(* IEC 61131-3 sources: PLC_I/plc/src/hardware, 9 files *)

(* ---- 全局变量_气缸IO映像.gvl.st ---- *)
(* 气缸物理 IO 映像。设备树把扩展输入/输出模块映射到本数组后，
   由 程序_气缸输入映射 / 程序_气缸输出映射 按工程表地址读写。
   容量：输入 112 点(7 WORD)，输出 56 点(4 WORD)。
   未映射时数组保持 0，模块在线位保持 FALSE，气缸许可因此关闭。 *)
VAR_GLOBAL CONSTANT
    ui气缸输入点数 : UINT := 112;
    ui气缸输出点数 : UINT := 56;
END_VAR
VAR_GLOBAL
    aw气缸输入映像 : ARRAY[0..6] OF WORD;
    aw气缸输出映像 : ARRAY[0..3] OF WORD;
    (* 真实模块诊断：由设备树/总线诊断赋值，不得用工程常量冒充。 *)
    b气缸输入模块在线 : BOOL;
    b气缸输出模块在线 : BOOL;
END_VAR

(* ---- 全局变量_气缸工程.gvl.st ---- *)
(* 唯一气缸工程配置：一缸一行，读起来就是接线表。
   默认全部未绑定，不驱动任何现场输出。
   点号 = 端子号（当前少量气缸全接内建点，直连模式）：
     in动点 := 5 就是 X5，out动点 := 2 就是 Y2；
   实际接线在 全局变量_物理IO.gvl.st 与 程序_气缸输入映射/输出映射.st，
   本表点号用于 HMI 显示与配置校验，必须和接线表一致。
   扩展模块缸的点号从 32 起，由设备树映射到 aw气缸输入/输出映像。
   示例（接好线后把 已绑定 改为 TRUE，并按实际核对点号/阀型/确认方式）：
       双电控夹紧缸：
       (已绑定 := TRUE, e阀型 := Cy阀型.双线圈保持,
        out动点 := 2, out原点 := 3,
        e动点确认 := Cy确认.传感器, in动点 := 5,
        e原点确认 := Cy确认.传感器, in原点 := 6),
       原点用时间确认的缸：e原点确认 := Cy确认.延时，省略 in原点。
       只用时间确认的推料缸：
       (已绑定 := TRUE, e阀型 := Cy阀型.单线圈复位, out动点 := 2) *)
VAR_GLOBAL CONSTANT
    Cy气缸配置 : ARRAY[0..53] OF 结构体_Cy气缸配置 := [
        (* CY00：X5/X6 传感器，Y2/Y3 阀；双电控。模板，未绑定 *)
        (已绑定 := FALSE, e阀型 := Cy阀型.双线圈保持,
         out动点 := 2, out原点 := 3,
         e动点确认 := Cy确认.传感器, in动点 := 5,
         e原点确认 := Cy确认.传感器, in原点 := 6),
        (* CY01：X7 动点传感器，原点延时确认，Y6/Y7 阀。模板，未绑定 *)
        (已绑定 := FALSE, e阀型 := Cy阀型.双线圈保持,
         out动点 := 6, out原点 := 7,
         e动点确认 := Cy确认.传感器, in动点 := 7,
         e原点确认 := Cy确认.延时),
        52((已绑定 := FALSE))
    ];
END_VAR

(* ---- 全局变量_物理IO.gvl.st ---- *)
(* 物理输入/输出边界：全工程只有本文件出现物理地址。
   信捷 HSIO 实测映射（与 HSIO 配置页、SDFCfg0 软元件配置对应）：
     一般输入：X0..X7、X10..X13（八进制编号，无 X8/X9）；
     一般输出：Y2、Y3、Y6、Y7、Y10..Y13；
     轴0：脉冲 Y0 / 方向 Y4；轴1：脉冲 Y1 / 方向 Y5；轴2/轴3 当前未启用。
   少量气缸直连模板（全接内建点，按现场接线改名/改地址；本文件是唯一地址来源）：
     CY00：动点开关 X5、原点开关 X6、动点阀 Y2、原点阀 Y3
     CY01：动点开关 X7、原点侧不接传感器（用延时确认）、动点阀 Y6、原点阀 Y7
   直连绑定行在 程序_气缸输入映射.st / 程序_气缸输出映射.st 末尾；
   扩展模块仍走 aw气缸输入映像/aw气缸输出映像（点号从 32 起），由设备树映射。
   维护规则：
     1) %IX/%QX 与端子丝印不完全对应（X10 以后按八进制推），改线必须同步更新本文件、
        docs/硬件IO对照表.md 与现场接线图；
     2) 轴2/轴3 若启用，方向端口为 Y6/Y7，会与本文件的 Y6/Y7 一般输出冲突；
     3) 急停 X3 只保证不进入软件滤波链；硬件滤波由 HSIO/SDFCfg 配置决定，
        安全响应仍由现场急停回路保证，本程序不是安全 PLC。 *)
VAR_GLOBAL
    b启动按钮 AT %IX0.0 : BOOL;   (* X0 启动，高有效 *)
    b暂停按钮 AT %IX0.1 : BOOL;   (* X1 暂停，高有效 *)
    b复位按钮 AT %IX0.2 : BOOL;   (* X2 复位，高有效 *)
    b急停按钮 AT %IX0.3 : BOOL;   (* X3 急停常开，TRUE=按下，断线不可诊断 *)
    b备用输入 AT %IX0.4 : BOOL;   (* X4 备用，高有效 *)

    (* ===== CY00 双电控（模板，按现场接线改名）===== *)
    bCY00_动点传感器 AT %IX0.5 : BOOL;  (* X5 动点开关 *)
    bCY00_原点传感器 AT %IX0.6 : BOOL;  (* X6 原点开关 *)
    bCY00_动点阀 AT %QX0.2 : BOOL;      (* Y2 动点阀 *)
    bCY00_原点阀 AT %QX0.3 : BOOL;      (* Y3 原点阀 *)

    (* ===== CY01 双电控，原点用时间确认（模板）===== *)
    bCY01_动点传感器 AT %IX0.7 : BOOL;  (* X7 动点开关 *)
    bCY01_动点阀 AT %QX0.6 : BOOL;      (* Y6 动点阀 *)
    bCY01_原点阀 AT %QX0.7 : BOOL;      (* Y7 原点阀 *)
END_VAR

(* ---- 全局变量_硬件.gvl.st ---- *)
VAR_GLOBAL CONSTANT
    (* Protocol milli-units. These are provisional caps for bench bring-up:
       edit per drive/mechanics rating and re-download. 0 would block every
       parameter write, so never publish an all-zero array. *)
    audi额定速度 : ARRAY[0..15] OF UDINT := [16(1000000)];      (* 1000 mm/s *)
    audi额定加速度 : ARRAY[0..15] OF UDINT := [16(10000000)];   (* 10000 mm/s² *)
    audi额定减速度 : ARRAY[0..15] OF UDINT := [16(10000000)];
    audi额定停止减速度 : ARRAY[0..15] OF UDINT := [16(20000000)];
END_VAR
VAR_GLOBAL
    (* Pulse axes have no external Ready input. Their availability is derived
       from MC feedback; it does not prove that a pulse drive has power. *)
    ab正限位 : ARRAY[0..2] OF BOOL;
    ab负限位 : ARRAY[0..2] OF BOOL;
    (* Cylinder commissioning seam. Sensor inputs default FALSE until the IO image
       is mapped; valve demands are written to 全局变量_气缸IO映像 by the output map. *)
    ab气缸模块就绪 : ARRAY[0..53] OF BOOL; (* 由真实模块在线位推导，不可手工赋值 *)
    ab气缸映射有效 : ARRAY[0..53] OF BOOL; (* 由绑定、配置有效和地址容量推导 *)
    ab气缸动点传感器 : ARRAY[0..53] OF BOOL;
    ab气缸原点传感器 : ARRAY[0..53] OF BOOL;
    ab气缸动点输出 : ARRAY[0..53] OF BOOL;
    ab气缸原点输出 : ARRAY[0..53] OF BOOL;
END_VAR

(* ---- 全局变量_绑定.gvl.st ---- *)
(* Engineering binding, not proof of physical availability. *)
VAR_GLOBAL CONSTANT
    ui轴总数 : UINT := 16;
    ui气缸总数 : UINT := 54;
    ui点位池容量 : UINT := 120;
    w已绑定轴 : WORD := 16#0007;
    w绑定纪元 : WORD := 2;
    (* Slots 0/1/2: XJ_Axis0 / XJ_Axis1 / BusMotionAxis.
       Device-tree AXIS_REF_SM3 references must NOT be redeclared here.
       Slots 3..15 unbound; cylinder wiring unverified, all unbound.
       Do not replace unknown online/ready feedback with TRUE. *)
END_VAR
VAR_GLOBAL
    (* 由 程序_气缸绑定 每扫描从工程记录推导，不再手工维护位掩码。 *)
    lw已绑定气缸 : LWORD := 0;
END_VAR

(* ---- 全局变量_运行配置.gvl.st ---- *)
(* 现场运行配置。全部为工程常量，不允许经 Modbus 写入。
   这些开关对应原程序 全局变量_系统 中的同名工程开关，语义保持不变：
   任何一项在被现场核验前保持 FALSE / 安全侧默认值。 *)
VAR_GLOBAL CONSTANT
    (* 正式工艺 POU 接入并完成评审后才允许改为 TRUE。
       为 FALSE 时命令 2（整机启动）被拒绝为 12，与原程序
       “NOT b正式流程已接入 → 拒绝” 的既有约定一致。 *)
    b正式流程已接入 : BOOL := FALSE;

    (* 硬限位输入是否真实接线。未接线时禁止关闭软限位，
       否则轴在软硬限位都不生效的情况下仍可运动。 *)
    b硬限位已接线 : BOOL := FALSE;

    (* 气缸IO模块是否已按电气图接入并核验。未接入时气缸保持离线，
       避免“填了工程表就动”的误判。接入后置 TRUE。 *)
    b气缸IO已接入 : BOOL := FALSE;

    (* 模块在线诊断是否已接入。FALSE 时以 b气缸IO已接入 作为就绪依据；
       TRUE 时改由 b气缸输入模块在线 / b气缸输出模块在线 真实判定。 *)
    b气缸IO模块诊断已接入 : BOOL := FALSE;

    (* X0 启动 / X1 暂停 / X2 复位 的软件去抖时间，原程序为 20 ms。
       急停 X3 不进入本软件滤波链；HSIO/SDFCfg 的硬件滤波另算，
       安全响应仍由现场急停回路保证，本程序不是安全 PLC。 *)
    di输入滤波时间ms : DINT := 20;

    (* 输出映像容量。只发布已实测的 Y6/Y7 两路，不得按逻辑槽数推断。 *)
    ui物理输出点数 : UINT := 2;

    (* 暂停后恢复允许的位置偏差，单位与轴位置一致（0.001 工程单位）。
       超过该值不阻止恢复，但会在恢复后由本块下发回位定位。 *)
    di暂停恢复容差 : DINT := 30;

    (* 暂停后确认静止的时间，原程序为 300 ms。停稳后才抓拍快照，
       减速距离不计入偏离。 *)
    di暂停停稳ms : DINT := 300;
END_VAR

(* ---- 程序_气缸绑定.st ---- *)
(* 把 Cy 配置表换算成绑定掩码与协议配置。每扫描最先执行。
   一行配置决定：是否绑定、阀型、两侧点地址和确认方式。
   选 Cy确认.延时 的一侧不绑定输入，由动作计时完成。 *)
PROGRAM 程序_气缸绑定
VAR
    i : UINT;
    w类型 : WORD;
    w动点输出 : WORD;
    w原点输出 : WORD;
    w动点输入 : WORD;
    w原点输入 : WORD;
    lw绑定 : LWORD;
END_VAR

lw绑定 := 0;
FOR i := 0 TO 53 DO
    w类型 := 0;
    w动点输出 := WORD#16#FFFF;
    w原点输出 := WORD#16#FFFF;
    w动点输入 := WORD#16#FFFF;
    w原点输入 := WORD#16#FFFF;
    IF 全局变量_气缸工程.Cy气缸配置[i].已绑定 THEN
        lw绑定 := lw绑定 OR SHL(LWORD#1, i);
        CASE 全局变量_气缸工程.Cy气缸配置[i].e阀型 OF
            Cy阀型.双线圈保持: w类型 := 1;
            Cy阀型.真空吸附: w类型 := 2;
            Cy阀型.真空带破真空: w类型 := 3;
        ELSE
            w类型 := 0;
        END_CASE;
        w动点输出 := 全局变量_气缸工程.Cy气缸配置[i].out动点;
        IF (w类型 = 1) OR (w类型 = 3) THEN
            w原点输出 := 全局变量_气缸工程.Cy气缸配置[i].out原点;
        END_IF;
        IF 全局变量_气缸工程.Cy气缸配置[i].e动点确认 = Cy确认.传感器 THEN
            w动点输入 := 全局变量_气缸工程.Cy气缸配置[i].in动点;
        END_IF;
        IF 全局变量_气缸工程.Cy气缸配置[i].e原点确认 = Cy确认.传感器 THEN
            w原点输入 := 全局变量_气缸工程.Cy气缸配置[i].in原点;
        END_IF;
        IF 全局变量_气缸工程.Cy气缸配置[i].动点反相 THEN w类型 := w类型 OR WORD#16#0004; END_IF;
        IF 全局变量_气缸工程.Cy气缸配置[i].原点反相 THEN w类型 := w类型 OR WORD#16#0008; END_IF;
    END_IF;
    (* 工程值变化时清掉现场确认，要求重新确认后才能进入自动流程。 *)
    IF (全局变量_保持区.Store.aw气缸配置[i, 0] <> w类型)
        OR (全局变量_保持区.Store.aw气缸配置[i, 1] <> w动点输出)
        OR (全局变量_保持区.Store.aw气缸配置[i, 2] <> w原点输出)
        OR (全局变量_保持区.Store.aw气缸配置[i, 3] <> w动点输入)
        OR (全局变量_保持区.Store.aw气缸配置[i, 4] <> w原点输入) THEN
        全局变量_保持区.Store.b已确认 := FALSE;
    END_IF;
    全局变量_保持区.Store.aw气缸配置[i, 0] := w类型;
    全局变量_保持区.Store.aw气缸配置[i, 1] := w动点输出;
    全局变量_保持区.Store.aw气缸配置[i, 2] := w原点输出;
    全局变量_保持区.Store.aw气缸配置[i, 3] := w动点输入;
    全局变量_保持区.Store.aw气缸配置[i, 4] := w原点输入;
END_FOR;
全局变量_绑定.lw已绑定气缸 := lw绑定;
END_PROGRAM

(* ---- 程序_气缸输入映射.st ---- *)
(* 气缸输入映射：把物理输入换算成逻辑端位传感器，并推导"映射有效/模块就绪"。
   必须在 气缸调度 之前调用。本 POU 不产生任何输出驱动。
   两种来源：
     1) 扩展模块：按工程表点号从 aw气缸输入映像 读取（点号从 32 起）；
     2) 直连模式：少量气缸全接内建点，命名 BOOL 直接覆盖（见文件末尾）。 *)
PROGRAM 程序_气缸输入映射
VAR
    i : UINT;
    ui地址 : UINT;
    b模块就绪 : BOOL;
END_VAR

IF 全局变量_运行配置.b气缸IO模块诊断已接入 THEN
    b模块就绪 := b气缸输入模块在线 AND b气缸输出模块在线;
ELSE
    b模块就绪 := 全局变量_运行配置.b气缸IO已接入;
END_IF;

FOR i := 0 TO 53 DO
    ab气缸动点传感器[i] := FALSE;
    ab气缸原点传感器[i] := FALSE;
    ab气缸映射有效[i] := FALSE;
    IF (lw已绑定气缸 AND SHL(LWORD#1, i)) <> 0 THEN
        ab气缸映射有效[i] := 气缸_配置有效(缸号 := i, Store := 全局变量_保持区.Store);
        IF ab气缸映射有效[i] THEN
            ui地址 := WORD_TO_UINT(全局变量_保持区.Store.aw气缸配置[i, 3]);
            IF (ui地址 <> 65535) AND (ui地址 < ui气缸输入点数) THEN
                ab气缸动点传感器[i] :=
                    (aw气缸输入映像[ui地址 / 16] AND SHL(WORD#1, ui地址 MOD 16)) <> 0;
            END_IF;
            ui地址 := WORD_TO_UINT(全局变量_保持区.Store.aw气缸配置[i, 4]);
            IF (ui地址 <> 65535) AND (ui地址 < ui气缸输入点数) THEN
                ab气缸原点传感器[i] :=
                    (aw气缸输入映像[ui地址 / 16] AND SHL(WORD#1, ui地址 MOD 16)) <> 0;
            END_IF;
        END_IF;
    END_IF;
    ab气缸模块就绪[i] := b模块就绪;
END_FOR;

(* ===== 直连模式：命名传感器 -> 驱动数组 =====
   加直连缸时在此加对应行，并同步 程序_气缸输出映射 与 全局变量_气缸工程。 *)
ab气缸动点传感器[0] := bCY00_动点传感器;
ab气缸原点传感器[0] := bCY00_原点传感器;
ab气缸动点传感器[1] := bCY01_动点传感器;
END_PROGRAM

(* ---- 程序_气缸输出映射.st ---- *)
(* 气缸输出映射：把调度产生的逻辑阀需求写到物理输出。
   必须在 气缸调度 之后调用。两种去向：
     1) 扩展模块：按工程表点号写 aw气缸输出映像（点号从 32 起）；
     2) 直连模式：少量气缸全接内建点，直接驱动命名阀（见文件末尾）。 *)
PROGRAM 程序_气缸输出映射
VAR
    i : UINT;
    ui地址 : UINT;
END_VAR

FOR i := 0 TO 3 DO
    aw气缸输出映像[i] := 0;
END_FOR;
FOR i := 0 TO 53 DO
    IF (lw已绑定气缸 AND SHL(LWORD#1, i)) <> 0
        AND ab气缸映射有效[i] AND ab气缸模块就绪[i] THEN
        ui地址 := WORD_TO_UINT(全局变量_保持区.Store.aw气缸配置[i, 1]);
        IF (ui地址 <> 65535) AND (ui地址 < ui气缸输出点数)
            AND ab气缸动点输出[i] THEN
            aw气缸输出映像[ui地址 / 16] :=
                aw气缸输出映像[ui地址 / 16] OR SHL(WORD#1, ui地址 MOD 16);
        END_IF;
        ui地址 := WORD_TO_UINT(全局变量_保持区.Store.aw气缸配置[i, 2]);
        IF (ui地址 <> 65535) AND (ui地址 < ui气缸输出点数)
            AND ab气缸原点输出[i] THEN
            aw气缸输出映像[ui地址 / 16] :=
                aw气缸输出映像[ui地址 / 16] OR SHL(WORD#1, ui地址 MOD 16);
        END_IF;
    END_IF;
END_FOR;

(* ===== 直连模式：驱动数组 -> 命名阀（Y2/Y3/Y6/Y7）=====
   未绑定或映射无效时数组为 FALSE，阀输出为 0。加直连缸时在此加对应行。 *)
bCY00_动点阀 := ab气缸动点输出[0];
bCY00_原点阀 := ab气缸原点输出[0];
bCY01_动点阀 := ab气缸动点输出[1];
bCY01_原点阀 := ab气缸原点输出[1];
END_PROGRAM
